(* IEC 61131-3 sources: test/Class/SafetyBaseFSoE (part 3) *)

                // get length of Name
                sd_retval := SDOReadCfgRequ ( p_SDORequestBuffer  := p_SDORequestBuffer
                                            , p_SDOResponseBuffer := p_SDOResponseBuffer
                                            , ud_Address          := ud_Address
                                            , us_Length           := 4
                                            );
                //no response
                if ( sd_retval <> 0 ) then
                  LogError("@020A (SafetyBaseFSoE::ReadSDOConfig) Config Read Error: Reading length of unsafe BDINT output name failed.");
                  return;
                end_if;

                // prepare address to get name
                ud_Address += 4;

  //              ud_ActStrLen := ud_TmpStrLen := p_SDOResponseBuffer^.ud_Data;
                ud_TmpStrLen := p_SDOResponseBuffer^.ud_Data;
                ud_ActStrLen := ud_TmpStrLen;
                ud_TmpAddress := ud_Address;

                IF p_BlockedTransferMemory = NIL THEN
                  sd_retval := -100;
                  SetSafetyState(NewState:=_MemAllocFailed);
                  RETURN;
                END_IF;

                IF ud_BlockedTransferMemorySize < (ud_TmpStrLen + 1) THEN
                  p_BlockedTransferMemory := ToStdLib.ReAlloc(mptr:=p_BlockedTransferMemory, newsize:=GetNewMemSize(ud_TmpStrLen + 1));
                  IF p_BlockedTransferMemory = NIL THEN
                    ud_BlockedTransferMemorySize := 0;
                    sd_retval := -100;
                    SetSafetyState(NewState:=_MemAllocFailed);
                    RETURN;
                  ELSE
                    ud_BlockedTransferMemorySize := GetNewMemSize(ud_TmpStrLen + 1);
                  END_IF;
                END_IF;

                ToStdLib.MemSet(dest:=p_BlockedTransferMemory, value:=0, size:=ud_BlockedTransferMemorySize);

                p_TmpBlockedData := p_BlockedTransferMemory;

                us_BlockedTransferLength := BlockedTransferLength(ud_Datalength:=ud_TmpStrLen, us_MaxBlocklength:=60);

                while us_BlockedTransferLength do

                  // get name
                  sd_retval := SDOReadCfgRequ ( p_SDORequestBuffer  := p_SDORequestBuffer
                                              , p_SDOResponseBuffer := p_SDOResponseBuffer
                                              , ud_Address          := ud_TmpAddress
                                              , us_Length           := us_BlockedTransferLength
                                              , b_UseCache          := us_BlockedTransferLength < us_DataLength_Max
                                              );
                  //no response
                  if ( sd_retval <> 0 ) then
                    LogError("@0207 (SafetyBaseFSoE::ReadSDOConfig) Config Read Error: Reading unsafe BDINT output name failed.");
                    return;
                  end_if;

                  ToStdLib.MemCpy(dest:=p_TmpBlockedData,
                                   source:=#p_SDOResponseBuffer^.ud_Data,
                                   size:=us_BlockedTransferLength);

                  p_TmpBlockedData += us_BlockedTransferLength;
                  ud_TmpAddress += us_BlockedTransferLength;
                  ud_TmpStrLen -= us_BlockedTransferLength;

                  us_BlockedTransferLength := BlockedTransferLength(ud_Datalength:=ud_TmpStrLen, us_MaxBlocklength:=60);

                end_while;

                ActBitMask := (pBitMasks + (i-1) * sizeof(BDINT))^;

                // if unsafe component not found (sd_retval <> 0), it's not problem for whole safe application

                sd_retval :=AddFastUnsafeRoutElement(pRoutTable:=#p_FastUnsafeOutputsTable,
                                                     pRoutElementsNo:=#ui_CntFastUnsafeOutputs,
                                                     ud_Address:=ud_FastUnsafe_Offset_Out,
                                                     ui_NameLen:=ud_ActStrLen$UINT,
                                                     pNameNewElement:=p_BlockedTransferMemory$^CHAR,
                                                     ActBitMask,
                                                     bWriteVar:=TRUE);

                // get offset in application memory
                ud_ActAddress += CountBits(ActBitMask) * sizeof(DINT);
                ud_FastUnsafe_Offset_Out += sizeof(DINT);

                // prepare address for next unsafe output or for number of safe inputs
                ud_Address += ud_ActStrLen;

              end_for;

              // free the bitmasks
              ToStdLib.Free(mptr:=pBitMasks);

            end_if;

          end_if; //b_IprCodeLengthAvailable = FALSE

        end_if; //b_CfgTypeV2

//*****************************************************************************
//**   UNSAFE BOOL OUTPUT VARIABLES                                          **
//*****************************************************************************

        //read number of unsafe output vars

        //send request and receive data
        sd_retval := SDOReadCfgRequ ( p_SDORequestBuffer  := p_SDORequestBuffer
                                    , p_SDOResponseBuffer := p_SDOResponseBuffer
                                    , ud_Address          := ud_Address
                                    , us_Length           := 4
                                    );

        //no response
        if ( sd_retval <> 0 ) then
          LogError("@0204 (SafetyBaseFSoE::ReadSDOConfig) Config Read Error: Reading number of unsafe bool output vars failed.");
          return;
        end_if;

        ud_CntUnsafeOutputs := p_SDOResponseBuffer^.ud_Data;

        ud_Address += 4;

        // skip the names of unsafe outputs
        for i := 1 to ud_CntUnsafeOutputs do

          // get length of Name
          sd_retval := SDOReadCfgRequ ( p_SDORequestBuffer  := p_SDORequestBuffer
                                      , p_SDOResponseBuffer := p_SDOResponseBuffer
                                      , ud_Address          := ud_Address
                                      , us_Length           := 4
                                      );
          //no response
          if ( sd_retval <> 0 ) then
            LogError("@0205 (SafetyBaseFSoE::ReadSDOConfig) Config Read Error: Reading length of unsafe bool output name failed.");
            return;
          end_if;

          // prepare address to get name
          ud_Address += 4;

//          ud_ActStrLen := ud_TmpStrLen := p_SDOResponseBuffer^.ud_Data;
          ud_TmpStrLen := p_SDOResponseBuffer^.ud_Data;
          ud_ActStrLen := ud_TmpStrLen;
          ud_TmpAddress := ud_Address;

          IF p_BlockedTransferMemory = NIL THEN
            sd_retval := -100;
            SetSafetyState(NewState:=_MemAllocFailed);
            RETURN;
          END_IF;

          IF ud_BlockedTransferMemorySize < (ud_TmpStrLen + 1) THEN
            p_BlockedTransferMemory := ToStdLib.ReAlloc(mptr:=p_BlockedTransferMemory, newsize:=GetNewMemSize(ud_TmpStrLen + 1));
            IF p_BlockedTransferMemory = NIL THEN
              ud_BlockedTransferMemorySize := 0;
              sd_retval := -100;
              SetSafetyState(NewState:=_MemAllocFailed);
              RETURN;
            ELSE
              ud_BlockedTransferMemorySize := GetNewMemSize(ud_TmpStrLen + 1);
            END_IF;
          END_IF;

          ToStdLib.MemSet(dest:=p_BlockedTransferMemory, value:=0, size:=ud_BlockedTransferMemorySize);

          p_TmpBlockedData := p_BlockedTransferMemory;

          us_BlockedTransferLength := BlockedTransferLength(ud_Datalength:=ud_TmpStrLen, us_MaxBlocklength:=60);

          while us_BlockedTransferLength do

            // get name
            sd_retval := SDOReadCfgRequ ( p_SDORequestBuffer  := p_SDORequestBuffer
                                        , p_SDOResponseBuffer := p_SDOResponseBuffer
                                        , ud_Address          := ud_TmpAddress
                                        , us_Length           := us_BlockedTransferLength
                                        , b_UseCache          := us_BlockedTransferLength < us_DataLength_Max
                                        );
            //no response
            if ( sd_retval <> 0 ) then
              LogError("0206 (SafetyBaseFSoE::ReadSDOConfig) Config Read Error: Reading unsafe bool output name failed.");
              return;
            end_if;

            ToStdLib.MemCpy(dest:=p_TmpBlockedData,
                             source:=#p_SDOResponseBuffer^.ud_Data,
                             size:=us_BlockedTransferLength);

            p_TmpBlockedData += us_BlockedTransferLength;
            ud_TmpAddress += us_BlockedTransferLength;
            ud_TmpStrLen -= us_BlockedTransferLength;

            us_BlockedTransferLength := BlockedTransferLength(ud_Datalength:=ud_TmpStrLen, us_MaxBlocklength:=60);

          end_while;

          sd_retval := AddUnsafeRoutElement(pRoutTable:=#p_UnsafeOutputsTable,
                                            pRoutElementsNo:=#ui_CntUnsafeOutputs,
                                            ud_Address:=ud_ActAddress,
                                            ui_NameLen:=ud_ActStrLen$UINT,
                                            pNameNewElement:=p_BlockedTransferMemory$^CHAR);

          // if unsafe component not found (sd_retval <> 0), it's not problem for whole safe application

          // get offset in application memory
          ud_ActAddress += 4;

          // prepare address for next unsafe output or for number of safe inputs
          ud_Address += ud_ActStrLen;

        end_for;

        // special unsafe variables (not supported by old modules)
        if b_CfgTypeV2 then

//*****************************************************************************
//**   UNSAFE BDINT OUTPUT VARIABLES                                         **
//*****************************************************************************

          //read number of unsafe BDINT output vars

          //send request and receive data
          sd_retval := SDOReadCfgRequ ( p_SDORequestBuffer  := p_SDORequestBuffer
                                      , p_SDOResponseBuffer := p_SDOResponseBuffer
                                      , ud_Address          := ud_Address
                                      , us_Length           := 4
                                      );

          //no response
          if ( sd_retval <> 0 ) then
            LogError("@0207 (SafetyBaseFSoE::ReadSDOConfig) Config Read Error: Reading number of unsafe BDINT output vars failed.");
            return;
          end_if;

          ud_CntUnsafeOutputs := p_SDOResponseBuffer^.ud_Data;

          ud_Address += 4;

          if ud_CntUnsafeOutputs then

            //SDO request for this command has 5 bytes additional data
            pBitMasks$^void := ToStdLib.Malloc(size := ud_CntUnsafeOutputs * sizeof(BDINT));

            if ( pBitMasks = NIL ) then
              sd_retval                         := -100;
              SetSafetyState(NewState:=_MemAllocFailed);
              LogError("@0208 (SafetyBaseFSoE::ReadSDOConfig) Config Read Error: Failed to allocate memory for the BDINT variable bitmasks.");
              return;
            end_if;

            // get the bitmasks for the BDINT variables
            for i := 1 to ud_CntUnsafeOutputs do

              // get bitmask
              sd_retval := SDOReadCfgRequ ( p_SDORequestBuffer  := p_SDORequestBuffer
                                          , p_SDOResponseBuffer := p_SDOResponseBuffer
                                          , ud_Address          := ud_Address
                                          , us_Length           := 4
                                          );
              //no response
              if ( sd_retval <> 0 ) then
                LogError("@0207 (SafetyBaseFSoE::ReadSDOConfig) Config Read Error: Reading bit mask of unsafe BDINT output failed.");
                return;
              end_if;

              // prepare address for the next one
              ud_Address += 4;

              // save the bitmask for adding the rout element
              (pBitMasks + (i-1) * sizeof(BDINT))^ := p_SDOResponseBuffer^.ud_Data;
            end_for;

            // skip the names of unsafe outputs
            for i := 1 to ud_CntUnsafeOutputs do

              // get length of Name
              sd_retval := SDOReadCfgRequ ( p_SDORequestBuffer  := p_SDORequestBuffer
                                          , p_SDOResponseBuffer := p_SDOResponseBuffer
                                          , ud_Address          := ud_Address
                                          , us_Length           := 4
                                          );
              //no response
              if ( sd_retval <> 0 ) then
                LogError("@020A (SafetyBaseFSoE::ReadSDOConfig) Config Read Error: Reading length of unsafe BDINT output name failed.");
                return;
              end_if;

              // prepare address to get name
              ud_Address += 4;

//              ud_ActStrLen := ud_TmpStrLen := p_SDOResponseBuffer^.ud_Data;
              ud_TmpStrLen := p_SDOResponseBuffer^.ud_Data;
              ud_ActStrLen := ud_TmpStrLen;
              ud_TmpAddress := ud_Address;

              IF p_BlockedTransferMemory = NIL THEN
                sd_retval := -100;
                SetSafetyState(NewState:=_MemAllocFailed);
                RETURN;
              END_IF;

              IF ud_BlockedTransferMemorySize < (ud_TmpStrLen + 1) THEN
                p_BlockedTransferMemory := ToStdLib.ReAlloc(mptr:=p_BlockedTransferMemory, newsize:=GetNewMemSize(ud_TmpStrLen + 1));
                IF p_BlockedTransferMemory = NIL THEN
                  ud_BlockedTransferMemorySize := 0;
                  sd_retval := -100;
                  SetSafetyState(NewState:=_MemAllocFailed);
                  RETURN;
                ELSE
                  ud_BlockedTransferMemorySize := GetNewMemSize(ud_TmpStrLen + 1);
                END_IF;
              END_IF;

              ToStdLib.MemSet(dest:=p_BlockedTransferMemory, value:=0, size:=ud_BlockedTransferMemorySize);

              p_TmpBlockedData := p_BlockedTransferMemory;

              us_BlockedTransferLength := BlockedTransferLength(ud_Datalength:=ud_TmpStrLen, us_MaxBlocklength:=60);

              while us_BlockedTransferLength do

                // get name
                sd_retval := SDOReadCfgRequ ( p_SDORequestBuffer  := p_SDORequestBuffer
                                            , p_SDOResponseBuffer := p_SDOResponseBuffer
                                            , ud_Address          := ud_TmpAddress
                                            , us_Length           := us_BlockedTransferLength
                                            , b_UseCache          := us_BlockedTransferLength < us_DataLength_Max
                                            );
                //no response
                if ( sd_retval <> 0 ) then
                  LogError("@0207 (SafetyBaseFSoE::ReadSDOConfig) Config Read Error: Reading unsafe BDINT output name failed.");
                  return;
                end_if;

                ToStdLib.MemCpy(dest:=p_TmpBlockedData,
                                 source:=#p_SDOResponseBuffer^.ud_Data,
                                 size:=us_BlockedTransferLength);

                p_TmpBlockedData += us_BlockedTransferLength;
                ud_TmpAddress += us_BlockedTransferLength;
                ud_TmpStrLen -= us_BlockedTransferLength;

                us_BlockedTransferLength := BlockedTransferLength(ud_Datalength:=ud_TmpStrLen, us_MaxBlocklength:=60);

              end_while;

              ActBitMask := (pBitMasks + (i-1) * sizeof(BDINT))^;

              sd_retval := AddUnsafeRoutElement(pRoutTable:=#p_UnsafeOutputsTable,
                                                pRoutElementsNo:=#ui_CntUnsafeOutputs,
                                                ud_Address:=ud_UnsafeBDINT_Offset,
                                                ui_NameLen:=ud_ActStrLen$UINT,
                                                pNameNewElement:=p_BlockedTransferMemory$^CHAR,
                                                ActBitMask);

              // if unsafe component not found (sd_retval <> 0), it's not problem for whole safe application

              // get offset in application memory
              ud_ActAddress += CountBits(ActBitMask) * sizeof(DINT);
              ud_UnsafeBDINT_Offset += sizeof(DINT);

              // prepare address for next unsafe output or for number of safe inputs
              ud_Address += ud_ActStrLen;

            end_for;

            // free the bitmasks
            ToStdLib.Free(mptr:=pBitMasks);
          end_if;
        end_if;

//*****************************************************************************
//**   SAFE INPUT VARIABLES                                                  **
//*****************************************************************************

        // get number of safe inputs
        sd_retval := SDOReadCfgRequ ( p_SDORequestBuffer  := p_SDORequestBuffer
                                    , p_SDOResponseBuffer := p_SDOResponseBuffer
                                    , ud_Address          := ud_Address
                                    , us_Length           := 4
                                    );

        //no response
        if ( sd_retval <> 0 ) then
          LogError("@020B (SafetyBaseFSoE::ReadSDOConfig) Config Read Error: Reading number of safe inputs failed.");
          return;
        end_if;

        //number of safe inputs
        ud_TmpCnt := p_SDOResponseBuffer^.ud_Data;

        // get offset in application memory
        ud_ActAddress += ud_TmpCnt * 4;

        //address of path length of first safe input
        ud_Address := p_SDORequestBuffer^.ud_Address + 4;

        if ud_TmpCnt then
          //read path of all safe inputs and add them to routing lists
          for i := 1 to ud_TmpCnt do

            //read path
            sd_retval := ReadModulePath ( p_SDORequestBuffer          := p_SDORequestBuffer
                                        , p_SDOResponseBuffer         := p_SDOResponseBuffer
                                        , p_ud_Address                := #ud_Address
                                        , pModule                     := pModule
                                        , p_ud_ModulePathLen_Max      := #ud_ModulePathLen_Max
                                        , p_ud_ModulePathCompLen_Max  := #ud_ModulePathCompLen_Max
                                        , us_SDOMaxDataSize           := us_DataLength_Max
                                        );

            //no response, error
            if ( sd_retval <> 0 ) then
              LogError("@020C (SafetyBaseFSoE::ReadSDOConfig) Config Read Error: Reading path of safe input failed.");
              return;
            end_if;

            // if there is a valid module path
            if pModule^.p_us_Path <> NIL then
              //add module to routing tabs
              sd_retval := AddModuleToRoutingTabs ( pModule       := pModule
                                                  , pListHeader   := pListHeader
                                                  , b_IsOptional  := TempModuleConfig.Info.IsOptional
                                                  );

              if (sd_retval <> 0 ) then
                if ( SafetyState <> _ModFromCfgNotFound ) then
                  LogError("@020D (SafetyBaseFSoE::ReadSDOConfig) Config Read Error: Failed to add safe input module to routing tabs.");
                  return;
                end_if;
              end_if;
            end_if;

            if b_IsFSoE then
              // lower 2 Bytes: Index in connection list, upper 2 Bytes: Bit-Offset of the value inside the process data (not the FSoE frame)
              ud_Address += 4;
            else
              //address of path length = last address + 2 * 4 bytes ( RemoteIndex + MaxAge)
              ud_Address += 8;
            end_if;
          end_for;
        end_if;

        if b_CfgTypeV3 then

//*****************************************************************************
//**   SAFE DINT INPUT VARIABLES                                             **
//*****************************************************************************

          // get number of safe DINT inputs
          sd_retval := SDOReadCfgRequ ( p_SDORequestBuffer  := p_SDORequestBuffer
                                      , p_SDOResponseBuffer := p_SDOResponseBuffer
                                      , ud_Address          := ud_Address
                                      , us_Length           := 4
                                      );

          //no response
          if ( sd_retval <> 0 ) then
            LogError("@020E (SafetyBaseFSoE::ReadSDOConfig) Config Read Error: Reading number of safe DINT inputs failed.");
            return;
          end_if;

          //number of safe inputs
          ud_TmpCnt := p_SDOResponseBuffer^.ud_Data;

          // get offset in application memory
          ud_ActAddress += ud_TmpCnt * 8;

          //address of path length of first safe input
          ud_Address := p_SDORequestBuffer^.ud_Address + 4;

          //read path of all safe inputs and add them to routing lists
          for i := 1 to ud_TmpCnt do

            //read path
            sd_retval := ReadModulePath ( p_SDORequestBuffer          := p_SDORequestBuffer
                                        , p_SDOResponseBuffer         := p_SDOResponseBuffer
                                        , p_ud_Address                := #ud_Address
                                        , pModule                     := pModule
                                        , p_ud_ModulePathLen_Max      := #ud_ModulePathLen_Max
                                        , p_ud_ModulePathCompLen_Max  := #ud_ModulePathCompLen_Max
                                        , us_SDOMaxDataSize           := us_DataLength_Max
                                        );

            //no response, error
            if ( sd_retval <> 0 ) then
              LogError("@020F (SafetyBaseFSoE::ReadSDOConfig) Config Read Error: Reading path of safe DINT input failed.");
              return;
            end_if;

            // if there is a valid module path
            if pModule^.p_us_Path <> NIL then
              //add module to routing tabs
              sd_retval := AddModuleToRoutingTabs ( pModule       := pModule
                                                  , pListHeader   := pListHeader
                                                  , b_IsOptional  := TempModuleConfig.Info.IsOptional
                                                  );

              if (sd_retval <> 0 ) then
                if ( SafetyState <> _ModFromCfgNotFound ) then
                  LogError("@0210 (SafetyBaseFSoE::ReadSDOConfig) Config Read Error: Failed to add safe DINT input module to routing tabs.");
                  return;
                end_if;
              end_if;
            end_if;

            if b_IsFSoE then
              // lower 2 Bytes: Index in connection list, upper 2 Bytes: Bit-Offset of the value inside the process data (not the FSoE frame)
              ud_Address += 4;
            else
              //address of path length = last address + 2 * 4 bytes ( RemoteIndex + MaxAge)
              ud_Address += 8;
            end_if;
          end_for;
        end_if;

        // only available at new modules
        if b_CfgTypeV2 then

//*****************************************************************************
//**   SAFE INTERFACE INPUT VARIABLES                                        **
//*****************************************************************************

          // get number of safe interface input vars

          //send request and receive data
          sd_retval := SDOReadCfgRequ ( p_SDORequestBuffer  := p_SDORequestBuffer
                                      , p_SDOResponseBuffer := p_SDOResponseBuffer
                                      , ud_Address          := ud_Address
                                      , us_Length           := 4
                                      );

          //no response
          if ( sd_retval <> 0 ) then
            LogError("@0211 (SafetyBaseFSoE::ReadSDOConfig) Config Read Error: Reading number of safe interface input variables failed.");
            return;
          end_if;

          // skip the number
          ud_Address += 4;

          //number of safe inputs
          ud_TmpCnt := p_SDOResponseBuffer^.ud_Data;

          // get offset in application memory
          ud_ActAddress += ud_TmpCnt * 4;

          if ud_TmpCnt then

            for i := 0 to (ud_TmpCnt-1) do
              // get length of the uncompressed path

              //send request and receive data
              sd_retval := SDOReadCfgRequ ( p_SDORequestBuffer  := p_SDORequestBuffer
                                          , p_SDOResponseBuffer := p_SDOResponseBuffer
                                          , ud_Address          := ud_Address
                                          , us_Length           := 4
                                          );

              //no response
              if ( sd_retval <> 0 ) then
                LogError("@0212 (SafetyBaseFSoE::ReadSDOConfig) Config Read Error: Reading length of uncompressed interface topology path failed.");
                return;
              end_if;

              // skip length of top path
              ud_Address += 4;

              // skip top path
              ud_Address += p_SDOResponseBuffer^.ud_Data;

              // read length of compressed topology path

              //send request and receive data
              sd_retval := SDOReadCfgRequ ( p_SDORequestBuffer  := p_SDORequestBuffer
                                          , p_SDOResponseBuffer := p_SDOResponseBuffer
                                          , ud_Address          := ud_Address
                                          , us_Length           := 4
                                          );

              //no response
              if ( sd_retval <> 0 ) then
                LogError("@0279 (SafetyBaseFSoE::ReadSDOConfig) Config Read Error: Reading length of compressed interface topology path failed.");
                return;
              end_if;

              // skip length of compressed top path and compressed top path
              ud_Address += 4 + p_SDOResponseBuffer^.ud_Data;

              if b_IsFSoE then
                // lower 2 Bytes: Index in connection list, upper 2 Bytes: Bit-Offset of the value inside the process data (not the FSoE frame)
                ud_Address += 4;
              else
                //address of path length = last address + 2 * 4 bytes ( RemoteIndex + MaxAge)
                ud_Address += 8;
              end_if;
            end_for;
          end_if;

(*
 4 Byte Anzahl
 4 Byte Länge vom Pfad, Pfad (vorne Pfad ":" dann CRC für da Interface dann bis auf 4 Byte aufgefüllt)
 4 Byte Länge vom komprimierten Pfad, komprimierter Pfad (vorne Pfad ":" dann CRC für da Interface dann bis auf 4 Byte aufgefüllt)
 4 Byte RemoteIndex
 4 Byte Maximales Alter
*)

        end_if;

        // only available at new containers
        if b_CfgTypeV3 then

//*****************************************************************************
//**   SAFE DINT INTERFACE INPUT VARIABLES                                   **
//*****************************************************************************

          // get number of safe DINT interface input vars

          //send request and receive data
          sd_retval := SDOReadCfgRequ ( p_SDORequestBuffer  := p_SDORequestBuffer
                                      , p_SDOResponseBuffer := p_SDOResponseBuffer
                                      , ud_Address          := ud_Address
                                      , us_Length           := 4
                                      );

          //no response
          if ( sd_retval <> 0 ) then
            LogError("@0213 (SafetyBaseFSoE::ReadSDOConfig) Config Read Error: Reading number of safe DINT interface input variables failed.");
            return;
          end_if;

          // skip the number
          ud_Address += 4;

          //number of safe inputs
          ud_TmpCnt := p_SDOResponseBuffer^.ud_Data;

          // get offset in application memory
          ud_ActAddress += ud_TmpCnt * 8;

          if ud_TmpCnt then

            for i := 0 to (ud_TmpCnt-1) do
              // get length of the uncompressed path

              //send request and receive data
              sd_retval := SDOReadCfgRequ ( p_SDORequestBuffer  := p_SDORequestBuffer
                                          , p_SDOResponseBuffer := p_SDOResponseBuffer
                                          , ud_Address          := ud_Address
                                          , us_Length           := 4
                                          );

              //no response
              if ( sd_retval <> 0 ) then
                LogError("@0214 (SafetyBaseFSoE::ReadSDOConfig) Config Read Error: Reading length of uncompressed interface topology path failed at safe DINT input variables.");
                return;
              end_if;

              // skip length of top path
              ud_Address += 4;

              // skip top path
              ud_Address += p_SDOResponseBuffer^.ud_Data;

              // read length of compressed topology path

              //send request and receive data
              sd_retval := SDOReadCfgRequ ( p_SDORequestBuffer  := p_SDORequestBuffer
                                          , p_SDOResponseBuffer := p_SDOResponseBuffer
                                          , ud_Address          := ud_Address
                                          , us_Length           := 4
                                          );

              //no response
              if ( sd_retval <> 0 ) then
                LogError("@0215 (SafetyBaseFSoE::ReadSDOConfig) Config Read Error: Reading length of compressed interface topology path failed at safe DINT input variables.");
                return;
              end_if;

              // skip length of compressed top path and compressed top path
              ud_Address += 4 + p_SDOResponseBuffer^.ud_Data;

              if b_IsFSoE then
                // lower 2 Bytes: Index in connection list, upper 2 Bytes: Bit-Offset of the value inside the process data (not the FSoE frame)
                ud_Address += 4;
              else
                //address of path length = last address + 2 * 4 bytes ( RemoteIndex + MaxAge)
                ud_Address += 8;
              end_if;
            end_for;
          end_if;

(*
 4 Byte Anzahl
 4 Byte Länge vom Pfad, Pfad (vorne Pfad ":" dann CRC für da Interface dann bis auf 4 Byte aufgefüllt)
 4 Byte Länge vom komprimierten Pfad, komprimierter Pfad (vorne Pfad ":" dann CRC für da Interface dann bis auf 4 Byte aufgefüllt)
 4 Byte RemoteIndex
 4 Byte Maximales Alter
*)

        end_if;

//*****************************************************************************
//**   FAST UNSAFE INPUT VARIABLES                                           **
//*****************************************************************************

        // only available at new modules
        if b_CfgTypeV2 then

          if b_IprCodeLengthAvailable = FALSE then
            // get number of fast unsafe intput vars

            //send request and receive data
            sd_retval := SDOReadCfgRequ ( p_SDORequestBuffer  := p_SDORequestBuffer
                                        , p_SDOResponseBuffer := p_SDOResponseBuffer
                                        , ud_Address          := ud_Address
                                        , us_Length           := 4
                                        );

            //no response
            if ( sd_retval <> 0 ) then
              LogError("@0216 (SafetyBaseFSoE::ReadSDOConfig) Config Read Error: Reading number of fast unsafe intput vars failed.");
              return;
            end_if;

            ud_Address += 4;

            // get offset in application memory
            ud_ActAddress += p_SDOResponseBuffer^.ud_Data * 4;
            // if it's our own path, remember the fast unsafe settings
            if (PathOfThisCPU[0]$UINT = (pListHeader^.p_us_Path$^UINT)^) & (ToStdLib.MemCmp(#PathOfThisCPU[0], pListHeader^.p_us_Path, PathOfThisCPU[0]$UINT + 2) = 0) then
              if (p_SDOResponseBuffer^.ud_Data <> 0) then
                if ActivateFastUnsafeIOs then
                  b_FastUnsafeInputsActive := TRUE;
                else
                  // error => can't go on like this
                  LogError("@0202 (SafetyBaseFSoE::ReadSDOConfig) Number or size of module accesses increased with new safety project!");
                  LogError("@0203 (SafetyBaseFSoE::ReadSDOConfig) => Can't continue, because the new data is not covered by the actual accesses! Restart Application!");

                  b_NeedApplicationRestart := TRUE;
                end_if;
              end_if;
            end_if;
          else  //b_IprCodeLengthAvailable = FALSE

//*****************************************************************************
//**   Fast UNSAFE BOOL INPUT VARIABLES     SCP211                           **
//*****************************************************************************

            // here we go for unsafe bool input vars

            // get number of unsafe input vars
            sd_retval := SDOReadCfgRequ ( p_SDORequestBuffer  := p_SDORequestBuffer
                                        , p_SDOResponseBuffer := p_SDOResponseBuffer
                                        , ud_Address          := ud_Address
                                        , us_Length           := 4
                                        );

            //no response
            if ( sd_retval <> 0 ) then
              LogError("@0217 (SafetyBaseFSoE::ReadSDOConfig) Config Read Error: Failed to read number of unsafe input vars.");
              return;
            end_if;

            ud_CntFastUnsafeInputs:= p_SDOResponseBuffer^.ud_Data;

            ud_Address += 4;

            // skip the names of unsafe inputs
            for i := 1 to ud_CntFastUnsafeInputs do

              // get length of Name
              sd_retval := SDOReadCfgRequ ( p_SDORequestBuffer  := p_SDORequestBuffer
                                          , p_SDOResponseBuffer := p_SDOResponseBuffer
                                          , ud_Address          := ud_Address
                                          , us_Length           := 4
                                          );
              //no response
              if ( sd_retval <> 0 ) then
                LogError("@0218 (SafetyBaseFSoE::ReadSDOConfig) Config Read Error: Reading length of unsafe input name failed.");
                return;
              end_if;

              // prepare address to get name
              ud_Address += 4;

    //          ud_ActStrLen := ud_TmpStrLen := p_SDOResponseBuffer^.ud_Data;
              ud_TmpStrLen := p_SDOResponseBuffer^.ud_Data;
              ud_ActStrLen := ud_TmpStrLen;
              ud_TmpAddress := ud_Address;

              IF p_BlockedTransferMemory = NIL THEN
                sd_retval := -100;
                SetSafetyState(NewState:=_MemAllocFailed);
                RETURN;
              END_IF;

              IF ud_BlockedTransferMemorySize < (ud_TmpStrLen + 1) THEN
                p_BlockedTransferMemory := ToStdLib.ReAlloc(mptr:=p_BlockedTransferMemory, newsize:=GetNewMemSize(ud_TmpStrLen + 1));
                IF p_BlockedTransferMemory = NIL THEN
                  ud_BlockedTransferMemorySize := 0;
                  sd_retval := -100;
                  SetSafetyState(NewState:=_MemAllocFailed);
                  RETURN;
                ELSE
                  ud_BlockedTransferMemorySize := GetNewMemSize(ud_TmpStrLen + 1);
                END_IF;
              END_IF;

              ToStdLib.MemSet(dest:=p_BlockedTransferMemory, value:=0, size:=ud_BlockedTransferMemorySize);

              p_TmpBlockedData := p_BlockedTransferMemory;

              us_BlockedTransferLength := BlockedTransferLength(ud_Datalength:=ud_TmpStrLen, us_MaxBlocklength:=60);

              while us_BlockedTransferLength do

                // get name
                sd_retval := SDOReadCfgRequ ( p_SDORequestBuffer  := p_SDORequestBuffer
                                            , p_SDOResponseBuffer := p_SDOResponseBuffer
                                            , ud_Address          := ud_TmpAddress
                                            , us_Length           := us_BlockedTransferLength
                                            , b_UseCache          := us_BlockedTransferLength < us_DataLength_Max
                                            );
                //no response
                if ( sd_retval <> 0 ) then
                  LogError("@0219 (SafetyBaseFSoE::ReadSDOConfig) Config Read Error: Reading unsafe input name failed.");
                  return;
                end_if;

                ToStdLib.MemCpy(dest:=p_TmpBlockedData,
                                 source:=#p_SDOResponseBuffer^.ud_Data,
                                 size:=us_BlockedTransferLength);

                p_TmpBlockedData += us_BlockedTransferLength;
                ud_TmpAddress += us_BlockedTransferLength;
                ud_TmpStrLen -= us_BlockedTransferLength;

                us_BlockedTransferLength := BlockedTransferLength(ud_Datalength:=ud_TmpStrLen, us_MaxBlocklength:=60);

              end_while;

              sd_retval := AddFastUnsafeRoutElement(pRoutTable:=#p_FastUnsafeInputsTable,
                                                    pRoutElementsNo:=#ui_CntFastUnsafeInputs,
                                                    ud_Address:=ud_FastUnsafe_Offset_In,
                                                    ui_NameLen:=ud_ActStrLen$UINT,
                                                    pNameNewElement:=p_BlockedTransferMemory$^CHAR,
                                                    bWriteVar:=FALSE);

              // if unsafe component not found (sd_retval <> 0), it's not problem for whole safe application
              // get offset in application memory
              ud_ActAddress += 4;
              ud_FastUnsafe_Offset_In += sizeof(DINT);

              // prepare address for next unsafe input
              ud_Address += ud_ActStrLen;

            end_for;

//*****************************************************************************
//**  FAST UNSAFE BDINT INPUT VARIABLES       SCP211                         **
//*****************************************************************************

            // here we go for unsafe BDINT input vars

            // get number of unsafe input vars
            sd_retval := SDOReadCfgRequ ( p_SDORequestBuffer  := p_SDORequestBuffer
                                        , p_SDOResponseBuffer := p_SDOResponseBuffer
                                        , ud_Address          := ud_Address
                                        , us_Length           := 4
                                        );

            //no response
            if ( sd_retval <> 0 ) then
              LogError("@021A (SafetyBaseFSoE::ReadSDOConfig) Config Read Error: Failed to read number of unsafe BDINT input vars.");
              return;
            end_if;

            ud_CntFastUnsafeInputs := p_SDOResponseBuffer^.ud_Data;

            ud_Address += 4;

            if ud_CntFastUnsafeInputs then

              //SDO request for this command has 5 bytes additional data
              pBitMasks$^void := ToStdLib.Malloc(size := ud_CntFastUnsafeInputs * sizeof(BDINT));

              if ( pBitMasks = NIL ) then
                sd_retval                         := -100;
                SetSafetyState(NewState:=_MemAllocFailed);
                LogError("@021B (SafetyBaseFSoE::ReadSDOConfig) Config Read Error: Failed to allocate memory for the BDINT variable bitmasks.");
                return;
              end_if;

              // get the bitmasks for the BDINT variables
              for i := 1 to ud_CntFastUnsafeInputs do

                // get bitmask
                sd_retval := SDOReadCfgRequ ( p_SDORequestBuffer  := p_SDORequestBuffer
                                            , p_SDOResponseBuffer := p_SDOResponseBuffer
                                            , ud_Address          := ud_Address
                                            , us_Length           := 4
                                            );
                //no response
                if ( sd_retval <> 0 ) then
                  LogError("021C (SafetyBaseFSoE::ReadSDOConfig) Config Read Error: Reading bit mask of unsafe BDINT input failed.");
                  return;
                end_if;

                // prepare address for the next one
                ud_Address += 4;

                // save the bitmask for adding the rout element
                (pBitMasks + (i-1) * sizeof(BDINT))^ := p_SDOResponseBuffer^.ud_Data;
              end_for;

              // get the names of unsafe inputs
              for i := 1 to ud_CntFastUnsafeInputs do

                // get length of Name
                sd_retval := SDOReadCfgRequ ( p_SDORequestBuffer  := p_SDORequestBuffer
                                            , p_SDOResponseBuffer := p_SDOResponseBuffer
                                            , ud_Address          := ud_Address
                                            , us_Length           := 4
                                            );
                //no response
                if ( sd_retval <> 0 ) then
                  LogError("@021D (SafetyBaseFSoE::ReadSDOConfig) Config Read Error: Reading length of unsafe BDINT input name failed.");
                  return;
                end_if;

                // prepare address to get name
                ud_Address += 4;

  //              ud_ActStrLen := ud_TmpStrLen := p_SDOResponseBuffer^.ud_Data;
                ud_TmpStrLen := p_SDOResponseBuffer^.ud_Data;
                ud_ActStrLen := ud_TmpStrLen;
                ud_TmpAddress := ud_Address;

                IF p_BlockedTransferMemory = NIL THEN
                  sd_retval := -100;
                  SetSafetyState(NewState:=_MemAllocFailed);
                  RETURN;
                END_IF;

                IF ud_BlockedTransferMemorySize < (ud_TmpStrLen + 1) THEN
                  p_BlockedTransferMemory := ToStdLib.ReAlloc(mptr:=p_BlockedTransferMemory, newsize:=GetNewMemSize(ud_TmpStrLen + 1));
                  IF p_BlockedTransferMemory = NIL THEN
                    ud_BlockedTransferMemorySize := 0;
                    sd_retval := -100;
                    SetSafetyState(NewState:=_MemAllocFailed);
                    RETURN;
                  ELSE
                    ud_BlockedTransferMemorySize := GetNewMemSize(ud_TmpStrLen + 1);
                  END_IF;
                END_IF;

                ToStdLib.MemSet(dest:=p_BlockedTransferMemory, value:=0, size:=ud_BlockedTransferMemorySize);

                p_TmpBlockedData := p_BlockedTransferMemory;

                us_BlockedTransferLength := BlockedTransferLength(ud_Datalength:=ud_TmpStrLen, us_MaxBlocklength:=60);

                while us_BlockedTransferLength do

                  // get name
                  sd_retval := SDOReadCfgRequ ( p_SDORequestBuffer  := p_SDORequestBuffer
                                              , p_SDOResponseBuffer := p_SDOResponseBuffer
                                              , ud_Address          := ud_TmpAddress
                                              , us_Length           := us_BlockedTransferLength
                                              , b_UseCache          := us_BlockedTransferLength < us_DataLength_Max
                                              );
                  //no response
                  if ( sd_retval <> 0 ) then
                    LogError("@021E (SafetyBaseFSoE::ReadSDOConfig) Config Read Error: Reading unsafe BDINT input name failed.");
                    return;
                  end_if;

                  ToStdLib.MemCpy(dest:=p_TmpBlockedData,
                                   source:=#p_SDOResponseBuffer^.ud_Data,
                                   size:=us_BlockedTransferLength);

                  p_TmpBlockedData += us_BlockedTransferLength;
                  ud_TmpAddress += us_BlockedTransferLength;
                  ud_TmpStrLen -= us_BlockedTransferLength;

                  us_BlockedTransferLength := BlockedTransferLength(ud_Datalength:=ud_TmpStrLen, us_MaxBlocklength:=60);

                end_while;

                ActBitMask := (pBitMasks + (i-1) * sizeof(BDINT))^;

                sd_retval := AddFastUnsafeRoutElement(pRoutTable:=#p_FastUnsafeInputsTable,
                                                      pRoutElementsNo:=#ui_CntFastUnsafeInputs,
                                                      ud_Address:=ud_FastUnsafe_Offset_In,
                                                      ui_NameLen:=ud_ActStrLen$UINT,
                                                      pNameNewElement:=p_BlockedTransferMemory$^CHAR,
                                                      BitMask:=ActBitMask,
                                                      bWriteVar:= FALSE);

                // if unsafe component not found (sd_retval <> 0), it's not problem for whole safe application

                // get offset in application memory
                ud_ActAddress += CountBits(ActBitMask) * sizeof(DINT);
                ud_FastUnsafe_Offset_In += sizeof(DINT);

                // prepare address for next unsafe output or for number of constants
                ud_Address += ud_ActStrLen;

              end_for;

              // free the bitmasks
              ToStdLib.Free(mptr:=pBitMasks);

            end_if;
        end_if;
      end_if; //b_CfgTypeV2

//*****************************************************************************
//**   UNSAFE BOOL INPUT VARIABLES                                           **
//*****************************************************************************

        // here we go for unsafe bool input vars

        // get number of unsafe input vars
        sd_retval := SDOReadCfgRequ ( p_SDORequestBuffer  := p_SDORequestBuffer
                                    , p_SDOResponseBuffer := p_SDOResponseBuffer
                                    , ud_Address          := ud_Address
                                    , us_Length           := 4
                                    );

        //no response
        if ( sd_retval <> 0 ) then
          LogError("@0217 (SafetyBaseFSoE::ReadSDOConfig) Config Read Error: Failed to read number of unsafe input vars.");
          return;
        end_if;

        ud_CntUnsafeInputs := p_SDOResponseBuffer^.ud_Data;

        ud_Address += 4;

        // skip the names of unsafe inputs
        for i := 1 to ud_CntUnsafeInputs do

          // get length of Name
          sd_retval := SDOReadCfgRequ ( p_SDORequestBuffer  := p_SDORequestBuffer
                                      , p_SDOResponseBuffer := p_SDOResponseBuffer
                                      , ud_Address          := ud_Address
                                      , us_Length           := 4
                                      );
          //no response
          if ( sd_retval <> 0 ) then
            LogError("@0218 (SafetyBaseFSoE::ReadSDOConfig) Config Read Error: Reading length of unsafe input name failed.");
            return;
          end_if;

          // prepare address to get name
          ud_Address += 4;

//          ud_ActStrLen := ud_TmpStrLen := p_SDOResponseBuffer^.ud_Data;
          ud_TmpStrLen := p_SDOResponseBuffer^.ud_Data;
          ud_ActStrLen := ud_TmpStrLen;
          ud_TmpAddress := ud_Address;

          IF p_BlockedTransferMemory = NIL THEN
            sd_retval := -100;
            SetSafetyState(NewState:=_MemAllocFailed);
            RETURN;
          END_IF;

          IF ud_BlockedTransferMemorySize < (ud_TmpStrLen + 1) THEN
            p_BlockedTransferMemory := ToStdLib.ReAlloc(mptr:=p_BlockedTransferMemory, newsize:=GetNewMemSize(ud_TmpStrLen + 1));
            IF p_BlockedTransferMemory = NIL THEN
              ud_BlockedTransferMemorySize := 0;
              sd_retval := -100;
              SetSafetyState(NewState:=_MemAllocFailed);
              RETURN;
            ELSE
              ud_BlockedTransferMemorySize := GetNewMemSize(ud_TmpStrLen + 1);
            END_IF;
          END_IF;

          ToStdLib.MemSet(dest:=p_BlockedTransferMemory, value:=0, size:=ud_BlockedTransferMemorySize);

          p_TmpBlockedData := p_BlockedTransferMemory;

          us_BlockedTransferLength := BlockedTransferLength(ud_Datalength:=ud_TmpStrLen, us_MaxBlocklength:=60);

          while us_BlockedTransferLength do

            // get name
            sd_retval := SDOReadCfgRequ ( p_SDORequestBuffer  := p_SDORequestBuffer
                                        , p_SDOResponseBuffer := p_SDOResponseBuffer
                                        , ud_Address          := ud_TmpAddress
                                        , us_Length           := us_BlockedTransferLength
                                        , b_UseCache          := us_BlockedTransferLength < us_DataLength_Max
                                        );
            //no response
            if ( sd_retval <> 0 ) then
              LogError("@0219 (SafetyBaseFSoE::ReadSDOConfig) Config Read Error: Reading unsafe input name failed.");
              return;
            end_if;

            ToStdLib.MemCpy(dest:=p_TmpBlockedData,
                             source:=#p_SDOResponseBuffer^.ud_Data,
                             size:=us_BlockedTransferLength);

            p_TmpBlockedData += us_BlockedTransferLength;
            ud_TmpAddress += us_BlockedTransferLength;
            ud_TmpStrLen -= us_BlockedTransferLength;

            us_BlockedTransferLength := BlockedTransferLength(ud_Datalength:=ud_TmpStrLen, us_MaxBlocklength:=60);

          end_while;

          sd_retval := AddUnsafeRoutElement(pRoutTable:=#p_UnsafeInputsTable,
                                            pRoutElementsNo:=#ui_CntUnsafeInputs,
                                            ud_Address:=ud_ActAddress,
                                            ui_NameLen:=ud_ActStrLen$UINT,
                                            pNameNewElement:=p_BlockedTransferMemory$^CHAR);

          // if unsafe component not found (sd_retval <> 0), it's not problem for whole safe application

          // get offset in application memory
          ud_ActAddress += 4;

          // prepare address for next unsafe input
          ud_Address += ud_ActStrLen;

        end_for;

        // only available at new modules
        if b_CfgTypeV2 then

//*****************************************************************************
//**   UNSAFE BDINT INPUT VARIABLES                                          **
//*****************************************************************************

          // here we go for unsafe BDINT input vars

          // get number of unsafe input vars
          sd_retval := SDOReadCfgRequ ( p_SDORequestBuffer  := p_SDORequestBuffer
                                      , p_SDOResponseBuffer := p_SDOResponseBuffer
                                      , ud_Address          := ud_Address
                                      , us_Length           := 4
                                      );

          //no response
          if ( sd_retval <> 0 ) then
            LogError("@021A (SafetyBaseFSoE::ReadSDOConfig) Config Read Error: Failed to read number of unsafe BDINT input vars.");
            return;
          end_if;

          ud_CntUnsafeInputs := p_SDOResponseBuffer^.ud_Data;

          ud_Address += 4;

          if ud_CntUnsafeInputs then

            //SDO request for this command has 5 bytes additional data
            pBitMasks$^void := ToStdLib.Malloc(size := ud_CntUnsafeInputs * sizeof(BDINT));

            if ( pBitMasks = NIL ) then
              sd_retval                         := -100;
              SetSafetyState(NewState:=_MemAllocFailed);
              LogError("@021B (SafetyBaseFSoE::ReadSDOConfig) Config Read Error: Failed to allocate memory for the BDINT variable bitmasks.");
              return;
            end_if;

            // get the bitmasks for the BDINT variables
            for i := 1 to ud_CntUnsafeInputs do

              // get bitmask
              sd_retval := SDOReadCfgRequ ( p_SDORequestBuffer  := p_SDORequestBuffer
                                          , p_SDOResponseBuffer := p_SDOResponseBuffer
                                          , ud_Address          := ud_Address
                                          , us_Length           := 4
                                          );
              //no response
              if ( sd_retval <> 0 ) then
                LogError("021C (SafetyBaseFSoE::ReadSDOConfig) Config Read Error: Reading bit mask of unsafe BDINT input failed.");
                return;
              end_if;

              // prepare address for the next one
              ud_Address += 4;

              // save the bitmask for adding the rout element
              (pBitMasks + (i-1) * sizeof(BDINT))^ := p_SDOResponseBuffer^.ud_Data;
            end_for;

            // get the names of unsafe inputs
            for i := 1 to ud_CntUnsafeInputs do

              // get length of Name
              sd_retval := SDOReadCfgRequ ( p_SDORequestBuffer  := p_SDORequestBuffer
                                          , p_SDOResponseBuffer := p_SDOResponseBuffer
                                          , ud_Address          := ud_Address
                                          , us_Length           := 4
                                          );
              //no response
              if ( sd_retval <> 0 ) then
                LogError("@021D (SafetyBaseFSoE::ReadSDOConfig) Config Read Error: Reading length of unsafe BDINT input name failed.");
                return;
              end_if;

              // prepare address to get name
              ud_Address += 4;

//              ud_ActStrLen := ud_TmpStrLen := p_SDOResponseBuffer^.ud_Data;
              ud_TmpStrLen := p_SDOResponseBuffer^.ud_Data;
              ud_ActStrLen := ud_TmpStrLen;
              ud_TmpAddress := ud_Address;

              IF p_BlockedTransferMemory = NIL THEN
                sd_retval := -100;
                SetSafetyState(NewState:=_MemAllocFailed);
                RETURN;
              END_IF;

              IF ud_BlockedTransferMemorySize < (ud_TmpStrLen + 1) THEN
                p_BlockedTransferMemory := ToStdLib.ReAlloc(mptr:=p_BlockedTransferMemory, newsize:=GetNewMemSize(ud_TmpStrLen + 1));
                IF p_BlockedTransferMemory = NIL THEN
                  ud_BlockedTransferMemorySize := 0;
                  sd_retval := -100;
                  SetSafetyState(NewState:=_MemAllocFailed);
                  RETURN;
                ELSE
                  ud_BlockedTransferMemorySize := GetNewMemSize(ud_TmpStrLen + 1);
                END_IF;
              END_IF;

              ToStdLib.MemSet(dest:=p_BlockedTransferMemory, value:=0, size:=ud_BlockedTransferMemorySize);

              p_TmpBlockedData := p_BlockedTransferMemory;

              us_BlockedTransferLength := BlockedTransferLength(ud_Datalength:=ud_TmpStrLen, us_MaxBlocklength:=60);

              while us_BlockedTransferLength do

                // get name
                sd_retval := SDOReadCfgRequ ( p_SDORequestBuffer  := p_SDORequestBuffer
                                            , p_SDOResponseBuffer := p_SDOResponseBuffer
                                            , ud_Address          := ud_TmpAddress
                                            , us_Length           := us_BlockedTransferLength
                                            , b_UseCache          := us_BlockedTransferLength < us_DataLength_Max
                                            );
                //no response
                if ( sd_retval <> 0 ) then
                  LogError("@021E (SafetyBaseFSoE::ReadSDOConfig) Config Read Error: Reading unsafe BDINT input name failed.");
                  return;
                end_if;

                ToStdLib.MemCpy(dest:=p_TmpBlockedData,
                                 source:=#p_SDOResponseBuffer^.ud_Data,
                                 size:=us_BlockedTransferLength);

                p_TmpBlockedData += us_BlockedTransferLength;
                ud_TmpAddress += us_BlockedTransferLength;
                ud_TmpStrLen -= us_BlockedTransferLength;

                us_BlockedTransferLength := BlockedTransferLength(ud_Datalength:=ud_TmpStrLen, us_MaxBlocklength:=60);

              end_while;

              ActBitMask := (pBitMasks + (i-1) * sizeof(BDINT))^;

              sd_retval := AddUnsafeRoutElement(pRoutTable:=#p_UnsafeInputsTable,
                                                pRoutElementsNo:=#ui_CntUnsafeInputs,
                                                ud_Address:=ud_UnsafeBDINT_Offset,
                                                ui_NameLen:=ud_ActStrLen$UINT,
                                                pNameNewElement:=p_BlockedTransferMemory$^CHAR,
                                                ActBitMask);

              // if unsafe component not found (sd_retval <> 0), it's not problem for whole safe application

              // get offset in application memory
              ud_ActAddress += CountBits(ActBitMask) * sizeof(DINT);
              ud_UnsafeBDINT_Offset += sizeof(DINT);

              // prepare address for next unsafe output or for number of constants
              ud_Address += ud_ActStrLen;

            end_for;

            // free the bitmasks
            ToStdLib.Free(mptr:=pBitMasks);
          end_if;

//*****************************************************************************
//**   CONSTANTS                                                             **
//*****************************************************************************

          // constants

          //send request and receive data
          sd_retval := SDOReadCfgRequ ( p_SDORequestBuffer  := p_SDORequestBuffer
                                      , p_SDOResponseBuffer := p_SDOResponseBuffer
                                      , ud_Address          := ud_Address
                                      , us_Length           := 4
                                      );

          //no response
          if ( sd_retval <> 0 ) then
            LogError("@021F (SafetyBaseFSoE::ReadSDOConfig) Config Read Error: Reading number of constants failed.");
            return;
          end_if;

          // skip number of constants
          ud_Address += 4;

          // skip constants
          ud_Address += p_SDOResponseBuffer^.ud_Data * 4;

          if b_CfgTypeV3 then

//*****************************************************************************
//**   SAFE DINT CONSTANTS                                                   **
//*****************************************************************************

            // constants

            //send request and receive data
            sd_retval := SDOReadCfgRequ ( p_SDORequestBuffer  := p_SDORequestBuffer
                                        , p_SDOResponseBuffer := p_SDOResponseBuffer
                                        , ud_Address          := ud_Address
                                        , us_Length           := 4
                                        );

            //no response
            if ( sd_retval <> 0 ) then
              LogError("@0220 (SafetyBaseFSoE::ReadSDOConfig) Config Read Error: Reading number of safe DINT constants failed.");
              return;
            end_if;

            // skip number of safe dint constants
            ud_Address += 4;

            // skip constants (4 byte per safe DINT constant)
            ud_Address += p_SDOResponseBuffer^.ud_Data * 4;

          end_if;

//*****************************************************************************
//**   LOCAL OUTPUTS                                                         **
//*****************************************************************************

          // local outputs
          //send request and receive data
          sd_retval := SDOReadCfgRequ ( p_SDORequestBuffer  := p_SDORequestBuffer
                                      , p_SDOResponseBuffer := p_SDOResponseBuffer
                                      , ud_Address          := ud_Address
                                      , us_Length           := 4
                                      );

          //no response
          if ( sd_retval <> 0 ) then
            LogError("@0221 (SafetyBaseFSoE::ReadSDOConfig) Config Read Error: Reading number of local outputs failed.");
            return;
          end_if;

          // skip number of local outputs
          ud_Address += 4;

          // skip local outputs
          //++pr
          // only available at new modules
          if b_CfgTypeV2 then
            ud_Address += p_SDOResponseBuffer^.ud_Data * 8; // Used-Flag, Modulkennung(SDIAS)
          else
            ud_Address += p_SDOResponseBuffer^.ud_Data * 4; // Used-Flag
          end_if;

          if b_CfgTypeV3 then

//*****************************************************************************
//**   LOCAL DINT OUTPUTS                                                    **
//*****************************************************************************

            // local outputs
            //send request and receive data
            sd_retval := SDOReadCfgRequ ( p_SDORequestBuffer  := p_SDORequestBuffer
                                        , p_SDOResponseBuffer := p_SDOResponseBuffer
                                        , ud_Address          := ud_Address
                                        , us_Length           := 4
                                        );

            //no response
            if ( sd_retval <> 0 ) then
              LogError("@0222 (SafetyBaseFSoE::ReadSDOConfig) Config Read Error: Reading number of local outputs failed.");
              return;
            end_if;

            // skip number of local outputs
            ud_Address += 4;

            // skip local outputs
            //++pr
            // only available at new modules
            if b_CfgTypeV2 then
              ud_Address += p_SDOResponseBuffer^.ud_Data * 8; // Used-Flag, Modulkennung(SDIAS)
            else
              ud_Address += p_SDOResponseBuffer^.ud_Data * 4; // Used-Flag
            end_if;

          end_if;

//*****************************************************************************
//**   SAFE BOOL INTERFACE OUTPUT VARIABLES                                  **
//*****************************************************************************

          // safe bool interface output vars
          //send request and receive data
          sd_retval := SDOReadCfgRequ ( p_SDORequestBuffer  := p_SDORequestBuffer
                                      , p_SDOResponseBuffer := p_SDOResponseBuffer
                                      , ud_Address          := ud_Address
                                      , us_Length           := 4
                                      );

          //no response
          if ( sd_retval <> 0 ) then
            LogError("@0223 (SafetyBaseFSoE::ReadSDOConfig) Config Read Error: Reading number of safe BOOL interface output variables failed.");
            return;
          end_if;

          // skip safe BOOL interface output variables
          ud_Address += 4;

          // count the interface output variables
          BoolOuts := p_SDOResponseBuffer^.ud_Data;

          if b_IsFSoE then
            ud_TmpCnt := p_SDOResponseBuffer^.ud_Data;

            if ud_TmpCnt then
              for i := 1 to ud_TmpCnt do
                //send request and receive data
                sd_retval := SDOReadCfgRequ ( p_SDORequestBuffer  := p_SDORequestBuffer
                                            , p_SDOResponseBuffer := p_SDOResponseBuffer
                                            , ud_Address          := ud_Address
                                            , us_Length           := 4
                                            );

                //no response
                if ( sd_retval <> 0 ) then
                  LogError("@027A (SafetyBaseFSoE::ReadSDOConfig) Config Read Error: Reading number of FSoE connections for BOOL interface outputs failed.");
                  return;
                end_if;

                // skip number of entries and the entries
                ud_Address += 4 + 4 * p_SDOResponseBuffer^.ud_Data;
              end_for;
            end_if;
          end_if;

//*****************************************************************************
//**   SAFE DINT INTERFACE OUTPUT VARIABLES                                  **
//*****************************************************************************

          // safe dint interface output vars
          //send request and receive data
          sd_retval := SDOReadCfgRequ ( p_SDORequestBuffer  := p_SDORequestBuffer
                                      , p_SDOResponseBuffer := p_SDOResponseBuffer
                                      , ud_Address          := ud_Address
                                      , us_Length           := 4
                                      );

          //no response
          if ( sd_retval <> 0 ) then
            LogError("@0224 (SafetyBaseFSoE::ReadSDOConfig) Config Read Error: Reading number of safe DINT interface output variables failed.");
            return;
          end_if;

          // skip number of safe dint interface output vars
          ud_Address += 4;

          // count the interface output variables
          DintOuts := p_SDOResponseBuffer^.ud_Data;

          if b_IsFSoE then
            ud_TmpCnt := p_SDOResponseBuffer^.ud_Data;

            if ud_TmpCnt then
              for i := 1 to ud_TmpCnt do
                //send request and receive data
                sd_retval := SDOReadCfgRequ ( p_SDORequestBuffer  := p_SDORequestBuffer
                                            , p_SDOResponseBuffer := p_SDOResponseBuffer
                                            , ud_Address          := ud_Address
                                            , us_Length           := 4
                                            );

                //no response
                if ( sd_retval <> 0 ) then
                  LogError("@027B (SafetyBaseFSoE::ReadSDOConfig) Config Read Error: Reading number of FSoE connections for DINT interface outputs failed.");
                  return;
                end_if;

                // skip number of entries and the entries
                ud_Address += 4 + 4 * p_SDOResponseBuffer^.ud_Data;
              end_for;
            end_if;
          end_if;

//*****************************************************************************
//**   FSBs = Functional Safety Blocks                                       **
//*****************************************************************************

          ud_skipLength := 0;

          // skip FSBs! structure: CRC, Length.... until the length is 0
          repeat

            // skip CRC and length of FSB
            ud_Address += 4 + ud_skipLength;

            //send request and receive data
            sd_retval := SDOReadCfgRequ ( p_SDORequestBuffer  := p_SDORequestBuffer
                                        , p_SDOResponseBuffer := p_SDOResponseBuffer
                                        , ud_Address          := ud_Address
                                        , us_Length           := 4
                                        );

            //no response
            if ( sd_retval <> 0 ) then
              LogError("@0225 (SafetyBaseFSoE::ReadSDOConfig) Config Read Error: Reading length of FSB failed.");
              return;
            end_if;

            ud_skipLength := p_SDOResponseBuffer^.ud_Data;

          until ud_skipLength = 0 end_repeat;

          // skip length of block with 0 length
          ud_Address += 4;

          if b_CfgTypeV3 then

//*****************************************************************************
//**   DYNAMIC PARAMETERS (e.g. for SSI Module)                              **
//*****************************************************************************

// Version of Parameters is saved in hd_DynParaVersion
// if it's 16#0001, then we read out the number of parameters which will follow

// structure:
// number of parameters
// for every parameter: place, id, length (including the 4 byte for the length itself), data

            //send request and receive data
            sd_retval := SDOReadCfgRequ ( p_SDORequestBuffer  := p_SDORequestBuffer
                                        , p_SDOResponseBuffer := p_SDOResponseBuffer
                                        , ud_Address          := ud_Address
                                        , us_Length           := 4
                                        );

            //no response
            if ( sd_retval <> 0 ) then
              LogError("@0226 (SafetyBaseFSoE::ReadSDOConfig) Config Read Error: Reading number of dynamic parameters failed.");
              return;
            end_if;

            ud_TmpCnt := p_SDOResponseBuffer^.ud_Data;

            // skip number of parameters
            ud_Address += 4;

            if ud_TmpCnt then
              for i := 1 to ud_TmpCnt do
                //send request and receive data
                sd_retval := SDOReadCfgRequ ( p_SDORequestBuffer  := p_SDORequestBuffer
                                            , p_SDOResponseBuffer := p_SDOResponseBuffer
                                            , ud_Address          := ud_Address
                                            , us_Length           := sizeof(t_DynamicParameterHeader)
                                            );

                //no response
                if ( sd_retval <> 0 ) then
                  LogError("@0227 (SafetyBaseFSoE::ReadSDOConfig) Config Read Error: Reading header of dynamic parameter failed.");
                  return;
                end_if;

                DynamicParameterHeader := p_SDOResponseBuffer^.ud_Data$t_DynamicParameterHeader;

                AddressServiceDataSize := 0;

                // skip size of header
                ud_Address += sizeof(t_DynamicParameterHeader);

                // data for pdo length info:
                // this data is also mirrored to SBF_SDO_ADDRESS_SPECIAL_INFO

//                  Marked with Place = 1000
//
//                  (4 Byte Length)
//                   4 Byte Version (starting at 0)
//                   1 Byte Length Rd PDO
//                   1 Byte Length Rd PDO IF
//                   1 Byte Length Wr PDO
//                   1 Byte Number of write PDOs (without additional it would be 1), msb = fast unsafe active

                if (DynamicParameterHeader.Place = SBF_CONFIG_PDO_INFO_PLACE) & (DynamicParameterHeader.Length >= (sizeof(UDINT) + sizeof(t_PDOSizeInfo))) then
                  //send request and receive data
                  sd_retval := SDOReadCfgRequ ( p_SDORequestBuffer  := p_SDORequestBuffer
                                              , p_SDOResponseBuffer := p_SDOResponseBuffer
                                              , ud_Address          := ud_Address
                                              , us_Length           := sizeof(t_PDOSizeInfo)
                                              );

                  //no response
                  if ( sd_retval <> 0 ) then
                    LogError("@0228 (SafetyBaseFSoE::ReadSDOConfig) Config Read Error: Reading dynamic parameter for pdo size failed.");
                    return;
                  end_if;

                  ud_Address += sizeof(t_PDOSizeInfo);

                  AddressServiceDataSize := (ud_ListLength_Address + ud_ListLength) - ud_Address;

                  PdoSizeInfo := p_SDOResponseBuffer^.ud_Data$t_PDOSizeInfo;

                  //check version
                  if PdoSizeInfo.Version = 1 then
                    // if any sizes increased or we would need more DOs
                    if (PdoSizeInfo.PDORdLen > MyPDOReadSize)     |
                       (PdoSizeInfo.PDOWrLen > MyPDOWriteSize)    |
                       ((PdoSizeInfo.FastUnsafeAvailable <> 0) > ActivateFastUnsafeIOs) then

                      // error => can't go on like this
                      LogError("@0202 (SafetyBaseFSoE::ReadSDOConfig) Number or size of module accesses increased with new safety project!");
                      LogError("@0203 (SafetyBaseFSoE::ReadSDOConfig) => Can't continue, because the new data is not covered by the actual accesses! Restart Application!");

                      b_NeedApplicationRestart := TRUE;
                    end_if;
                  else
                    // new interpretercode version
                    PdoSizeInfoV2 := p_SDOResponseBuffer^.ud_Data$t_PDOSizeInfoV2;

                    if  (PdoSizeInfoV2.PDORdLen > MyPDOReadSize)                       |
                        (PdoSizeInfoV2.PDOWrLen > MyPDOWriteSize)                      |
                        (PdoSizeInfoV2.uiNumberFastUnsafeRdVar > uiNumberFastUnsafeRd) |
                        (PdoSizeInfoV2.uiNumberFastUnsafeWrVar > uiNumberFastUnsafeWr) then

                      // error => can't go on like this
                      LogError("@0202 (SafetyBaseFSoE::ReadSDOConfig) Number or size of module accesses increased with new safety project!");
                      LogError("@0203 (SafetyBaseFSoE::ReadSDOConfig) => Can't continue, because the new data is not covered by the actual accesses! Restart Application!");

                      b_NeedApplicationRestart := TRUE;
                    end_if;
                  end_if;

                  exit;
                end_if;

                // skip the parameter data (length of the length is also included)
                ud_Address += DynamicParameterHeader.Length - 4;
              end_for;

              if AddressServiceDataSize then
(*

  Data structure of address service data

  4 Byte Anzahl der MultiChannel
    Pro MultiChannel:
    4 Byte Anzahl der Verwendungen des Multichannel
    4 Byte Index des Gesamtergebnisses
    1 Byte Art der Verknüpfung (0 = UND)
    1 Byte Defaultbelegung des Werts
    2 Byte Reserved (für 4 Byte Alignment)
      Pro Verwendung (siehe erster Eintrag in den MultiChannelDaten):
      4 Byte FSoE Daten
  4 Byte Kommunikations-ID (Default 0)
  4 Byte Anzahl der Adressbereiche
    Pro Adressbereich:
    4 Byte Startadresse
    4 Byte Länge Adressbereich
  4 Byte Anzahl der Connection-ID-Bereiche
    Pro Bereich:
    4 Byte Startadresse
    4 Byte Länge Bereich

*)
                // get the number of multichannels
                sd_retval := SDOReadCfgRequ ( p_SDORequestBuffer  := p_SDORequestBuffer
                                            , p_SDOResponseBuffer := p_SDOResponseBuffer
                                            , ud_Address          := ud_Address
                                            , us_Length           := 4
                                            );

                //no response
                if ( sd_retval <> 0 ) then
                  LogError("@027C (SafetyBaseFSoE::ReadSDOConfig) Config Read Error: Reading address service data failed.");
                  return;
                end_if;

                ud_TmpCnt := p_SDOResponseBuffer^.ud_Data;

                // skip number of multichannels
                ud_Address += 4;

                if ud_TmpCnt then
                  for i := 1 to ud_TmpCnt do
                    // get the number of usages
                    sd_retval := SDOReadCfgRequ ( p_SDORequestBuffer  := p_SDORequestBuffer
                                                , p_SDOResponseBuffer := p_SDOResponseBuffer
                                                , ud_Address          := ud_Address
                                                , us_Length           := 4
                                                );

                    //no response
                    if ( sd_retval <> 0 ) then
                      LogError("@027C (SafetyBaseFSoE::ReadSDOConfig) Config Read Error: Reading address service data failed.");
                      return;
                    end_if;

                    // skip the rest of this multichannel
                    ud_Address += 12 + (p_SDOResponseBuffer^.ud_Data * 4);
                  end_for;
                end_if;

                // skip the communication ID
                ud_Address += 4;

                // read the number of address areas
                sd_retval := SDOReadCfgRequ ( p_SDORequestBuffer  := p_SDORequestBuffer
                                            , p_SDOResponseBuffer := p_SDOResponseBuffer
                                            , ud_Address          := ud_Address
                                            , us_Length           := 4
                                            );

                //no response
                if ( sd_retval <> 0 ) then
                  LogError("@027C (SafetyBaseFSoE::ReadSDOConfig) Config Read Error: Reading address service data failed.");
                  return;
                end_if;

                // if there are any => the module got an address service
                if p_SDOResponseBuffer^.ud_Data then
                  TempModuleConfig.Info.IsAddressService := TRUE;
                end_if;
              end_if;
            end_if;
          end_if;

          // if there are interface variables
          if BoolOuts | DintOuts then
            // calculate the length of the interface frame
            TempPdoConfig.PdoLen := CalcPDOLength(BoolOuts, DintOuts);

            TempPdoConfig.Info := 0;
            TempPdoConfig.Info.IsInterfacePDO := TRUE;
            TempPdoConfig.Info.IsOptional := (ud_ActBlockType = SBF_BLKTYPE_CFG_MODULE_OPTIONAL);

            // if it's a broadcast => mark it
            if (TempPath[0]$UINT = 2) & (TempPath[0]$HDINT = SBF_INTERFACE_FRAME_BROADCAST) then
              TempPdoConfig.Info.IFBroadCast := TRUE;
            end_if;

            // this is the source of the interface frame
            TempPdoConfig.SourcePathLen := pListHeader^.p_us_Path^$UINT + 2;
            TempPdoConfig.pSourcePath   := pListHeader^.p_us_Path;

            // and the destination
            TempPdoConfig.DestPathLen   := TempPath[0]$UINT + 2;
            TempPdoConfig.pDestPath     := #TempPath[0];

            // add the interface PDO to the list
//            AddPdoToCfg(TempPdoConfig);

            TempModuleConfig.Info.IsInterfaceSource := TRUE;
            TempModuleConfig.Info.IsInterfaceDest   := FALSE;
            TempModuleConfig.InterfaceCRC := TempPdoConfig.InterfaceCRC;
          else
            TempModuleConfig.Info.IsInterfaceSource := FALSE;
            TempModuleConfig.Info.IsInterfaceDest   := FALSE;
            TempModuleConfig.InterfaceCRC := 0;
          end_if;
        else
          TempModuleConfig.Info.IsInterfaceSource := FALSE;
          TempModuleConfig.Info.IsInterfaceDest   := FALSE;
          TempModuleConfig.InterfaceCRC := 0;
        end_if;

        // if it's our own path, remember the safety number
        if (PathOfThisCPU[0]$UINT = (pListHeader^.p_us_Path$^UINT)^) & (ToStdLib.MemCmp(#PathOfThisCPU[0], pListHeader^.p_us_Path, PathOfThisCPU[0]$UINT + 2) = 0) then
          TempModuleConfig.SafetyNbr := SafetyNumber;
          //safe config of scp modul (own path)
          SafeActModuleConfig(TempModuleConfig);
        else
          TempModuleConfig.SafetyNbr := 0;
        end_if;

        // only when there is a manager
        if pSafetyManagerThis then
          AddModuleToCfg(TempModuleConfig);
        end_if;

//**********************************************************************************************************************************************************
      SBF_BLKTYPE_OLD_MODE_FLAG: // flag fore FW to use old config-mode
        // we need the old TimeSync config-type
        NewConfigType := ConfigState_Old;

//**********************************************************************************************************************************************************
      SBF_BLKTYPE_CFG_XML: // configuration for uploading the project to the safetydesigner (network placement information, names of bits,...)
        // no useful information here for us

//**********************************************************************************************************************************************************
    else
      // skip it = do nothing
//      TRACE("Found unhandled Blocktype in configuration.");
//**********************************************************************************************************************************************************
    end_case;

    ud_ListBaseAddress := ud_ListLength_Address + ud_ListLength;
  end_while;

  if ( ( sd_retval = 0 ) & ( SafetyState = _ModFromCfgNotFound ) ) then
    sd_retval := -1;
  end_if;

END_FUNCTION

FUNCTION VIRTUAL SafetyBaseFSoE::SDOReadCfgRequ
  VAR_INPUT
    p_SDORequestBuffer 	: ^SafetyBaseFSoE::SDORequReadConfig;
    p_SDOResponseBuffer 	: ^SafetyBaseFSoE::SDORespReadConfig;
    ud_Address 	: UDINT;
    us_Length 	: USINT;
    b_UseCache 	: BOOL;(* := TRUE *)
  END_VAR
  VAR_OUTPUT
    sd_retval 	: DINT;
  END_VAR

  // check if we have the data in the cache
  if b_UseCache & IsInCache(ud_Address, us_Length) then
    // use it from the cache

    // the address may be used from outside this function
    p_SDORequestBuffer^.ud_Address := ud_Address;

    _memcpy(ptr1:=#p_SDOResponseBuffer^.ud_Data, ptr2:=#Cache[0] + (ud_Address - CachedAddr), cntr:=us_Length);

    // everything is fine
    sd_retval := 0;
  else

    //sequence number
    p_SDORequestBuffer^.StdHeader.SeqNr := us_CntSequNr;

    //increase counter for sequence number
    if us_CntSequNr < 16#7F then
      us_CntSequNr += 1;
    else
      us_CntSequNr := 0;
    end_if;

    //address
    p_SDORequestBuffer^.ud_Address := ud_Address;

    if b_UseCache then
      // get max size
      p_SDORequestBuffer^.us_Length := SBF_SDO_MAX_LENGTH - (sizeof(SDORespReadConfig) - sizeof(SDORespReadConfig.ud_Data));
    else
      //length of expected data
      p_SDORequestBuffer^.us_Length := us_Length;
    end_if;

    //calculate CRC (starting with length of data until the end of command)
    p_SDORequestBuffer^.StdHeader.CRC := 0;

    //send request
    sd_retval := SAFETY_iSendRequest( uiMaster    := 0
                                    , pucNode     := p_ObjectPath
                                    , uiInLength  := sizeof(SDORequReadConfig)
                                    , pucInput    := p_SDORequestBuffer$^USINT
                                    , uiOutLength := sizeof(SDORespReadConfig) - sizeof(SDORespReadConfig.ud_Data) + p_SDORequestBuffer^.us_Length
                                    , pucOutput   := p_SDOResponseBuffer$^USINT
                                    );

    //no response
    if ( sd_retval <> 0 ) then
      LogError("@0229 (SafetyBaseFSoE::SDOReadCfgRequ) SAFETY_iSendRequest failed.");

      // we remember to retry in a few seconds
      b_ReadConfigFailed := TRUE;
      return;
    end_if;

    //check sequence number to exclude a possible wrong response
    if ( p_SDORequestBuffer^.StdHeader.SeqNr <> p_SDOResponseBuffer^.StdHeader.SeqNr ) then
      // we remember to retry in a few seconds
      b_ReadConfigFailed := TRUE;
      //log not routable SDOs
      LogValue("@022A (SafetyBaseFSoE::SDOReadCfgRequ) Invalid Sequence number in SDO Standard Response. Got 0x{0} instead of expected 0x{1}", to_udint(p_SDOResponseBuffer^.StdHeader.SeqNr), to_udint(p_SDORequestBuffer^.StdHeader.SeqNr));
      return;
    end_if;

    //check returncode of SDO
    if ( p_SDOResponseBuffer^.us_Returncode <> SBF_SDO_RETCODE_OK ) then
      //log not routable SDOs
      LogValue("@022B (SafetyBaseFSoE::SDOReadCfgRequ) Safety module 0x{0}: Retcode of SDO Standard Response was invalid. Retcode: 0x{1}", SafetyNumber$UDINT, to_udint(p_SDOResponseBuffer^.us_Returncode));

  //    // when reading fails because safety designer is writing at the same moment
  //    if p_SDOResponseBuffer^.us_Returncode = SDO_MICROCTRL_DIFFER then
        // we remember to retry in a few seconds
        b_ReadConfigFailed := TRUE;
  //    end_if;

      return;
    end_if;

    //check length of read data
    if ( p_SDOResponseBuffer^.us_Length = 0 ) then
      LogError("@022C (SafetyBaseFSoE::SDOReadCfgRequ) Response length is 0.");
      sd_retval := -104;
      return;
    elsif b_UseCache then
      // everything is fine => add the new data to the cache
      AddToCache(p_SDORequestBuffer, p_SDOResponseBuffer);
    end_if;
  end_if;

END_FUNCTION

FUNCTION VIRTUAL SafetyBaseFSoE::GetRoutingData
  VAR_OUTPUT
    sd_retval 	: DINT;
  END_VAR
  VAR
    SDORequestBuffer        : SDORequReadConfig;
    SDOResponseBuffer       : ARRAY [0..SBF_SDO_MAX_LENGTH-1] OF USINT;
    p_SDORequestBuffer 	    : ^SDORequReadConfig;
    p_SDOResponseBuffer 	  : ^SDORespReadConfig;
    Module                  : PathInfoType;
    ListHeader              : PathInfoType;
    NotAvailableStr         : ARRAY [0..99] OF CHAR;
    ModulePath              : ARRAY [0..127] OF USINT;
    ModulePathComp          : ARRAY [0..127] OF USINT;
    ListPath                : ARRAY [0..127] OF USINT;
    ListPathComp            : ARRAY [0..127] OF USINT;
    Time1, Time2            : UDINT;
  END_VAR

  // get module specific configuration information
  GetConfiguration();

  InitPathInfo(#Module);
  InitPathInfo(#ListHeader);

  //SDO request for this command has 5 bytes additional to the header
  p_SDORequestBuffer := #SDORequestBuffer;

  //SDO response for this command can have maximum additional data
  p_SDOResponseBuffer := (#SDOResponseBuffer)$^SDORespReadConfig;

  //path of input-safety-module
  Module.p_us_Path$^void := #ModulePath;

  //compressed path of input-safety-module
  Module.p_us_PathComp$^void := #ModulePathComp;

  //path in list header
  ListHeader.p_us_Path$^void := #ListPath;

  //path in list header
  ListHeader.p_us_PathComp$^void := #ListPathComp;

  repeat
    // if not used => continue
    // if valid    => set to not used and continue
    // if wait4rt  => wait in the loop until the state changes to valid
  until (sigclib_atomic_cmpxchgU32(pValue:=#udConfigValid, cmpVal:=SBF_LOCKCFG_VALID, newVal:=SBF_LOCKCFG_NOT_USED) < SBF_LOCKCFG_WAIT4RT) end_repeat;

  b_ReadConfigFailed := FALSE;

  b_NeedApplicationRestart := FALSE;

  // if there is a revision in the configuration this variable changes to TRUE
  b_GotNewRevision := FALSE;

Time1 := OS_READMICROSEC();
  //read config data via SDOs and add safety modules to routing lists
  sd_retval := ReadSDOConfig( p_SDORequestBuffer      := p_SDORequestBuffer
                            , p_SDOResponseBuffer     := p_SDOResponseBuffer
                            , pModule                 := #Module
                            , pListHeader             := #ListHeader
                            );
Time2 := OS_READMICROSEC();
ud_ConfigReadTime := Time2 - Time1;

  // set error to restart application afterwards to have a complete configuration (needed for routing to share the slave configurations with only 1 restart of the application)
  if b_NeedApplicationRestart then
    SetSafetyState(NewState:=_DOsIncreasedRestartApp);
    b_GetNewConfiguration := FALSE; // don't try again (unless the CRC changes again)
    sd_retval := -1;
  end_if;

  // if there is no revision in the configuration => clear it
  if (b_GotNewRevision = FALSE) then

    // free memory, if available
    if pPrjNameStr & pPrjRevStr then
      ToStdLib.Free(pPrjNameStr);
    end_if;

    // use local memory to show "not available"
    _strcpy(dest:=#NotAvailableStr[0], src:="<not available>");
    PrjNameMemLen := _strlen(src:=#NotAvailableStr[0]);
    PrjNameStrLen := PrjRevStrLen := PrjNameMemLen - 1;
    pPrjNameStr := pPrjRevStr := #NotAvailableStr[0];

    // write the strings to the string objects
    ShowProjectRevision();

    // there is no memory, so reset the pointer and length informations
    pPrjNameStr := NIL;
    pPrjRevStr := NIL;

    PrjNameMemLen := 0;
    PrjNameStrLen := 0;
    PrjRevStrLen := 0;
  end_if;

  // if reading failed, because designer is writing at the same time => we try again in a few seconds
  if b_ReadConfigFailed then

    // next time we check for the configured state of the cpu
    b_CheckConfigured := TRUE;
    b_GetNewConfiguration := FALSE; // don't try again while the config is invalid

    // check again in background
    SetSafetyState(NewState:=_ReinitConfig);

    // and wait at least 3 secs
    ud_LastCheckConfig := ops.tAbsolute;

  // error in configuration -> no work
  elsif ( sd_retval <> 0 ) & (SafetyState <> _ReinitConfig) then
    if SafetyState = _WaitForSynchronicity then
      SetSafetyState(NewState:=_UnknownCfgError);
    end_if;

    LogError("@022D (SafetyBaseFSoE::GetRoutingData) Reading Safety Configuration failed!");
  else
    // read config succeeded, check update cycle of unsafe variables
    CheckUnsafeUpdateCycle();

    // check for interface frame destination modules and mark them
    GetDestinationCRCs();

    // if there is a safety manager create a configuration message and send it to the safety manager
    if pSafetyManagerThis then
      CreateAndSendCfg();
    end_if;

    // last thing to do is to start realtime and cyclic work (they do nothing in _ReinitConfig state)
    if ud_UnsafeVarsNotFound then
      SetSafetyState(NewState:=_UnsafeVarNotFound);
      ud_UnsafeVarsNotFound := 0;
    else
      if us_SetBusReadyState = SetBusReadyFinished then
        // we're already synchron from a former configuration phase
        SetSafetyState(NewState:=_SafetyClassOK);
      else
        SetSafetyState(NewState:=_WaitForSynchronicity);
      end_if;
    end_if;

    // set config valid
    sigclib_atomic_swpU32(pValue:=#udConfigValid, swpVal:=SBF_LOCKCFG_VALID);
  end_if;

  // free temporary configuration lists if there were any
  FreeCfgLists();

END_FUNCTION

FUNCTION VIRTUAL SafetyBaseFSoE::ReadModulePath
  VAR_INPUT
    p_SDORequestBuffer 	: ^SafetyBaseFSoE::SDORequReadConfig;
    p_SDOResponseBuffer 	: ^SafetyBaseFSoE::SDORespReadConfig;
    p_ud_Address 	: ^UDINT;
    pModule 	: ^SafetyBaseFSoE::PathInfoType;
    p_ud_ModulePathLen_Max 	: ^UDINT;
    p_ud_ModulePathCompLen_Max 	: ^UDINT;
    us_SDOMaxDataSize 	: USINT;
  END_VAR
  VAR_OUTPUT
    sd_retval 	: DINT;
  END_VAR
  VAR
    ud_ModulePathLen_Act    : UDINT;
    p_ud_ModulePath_Act     : ^UDINT;
  END_VAR

  //read length of module path

  //send request and receive data
  sd_retval := SDOReadCfgRequ ( p_SDORequestBuffer  := p_SDORequestBuffer
                              , p_SDOResponseBuffer := p_SDOResponseBuffer
                              , ud_Address          := p_ud_Address^
                              , us_Length           := 4
                              );

  //no response
  if ( sd_retval <> 0 ) then
    LogError("@022E (SafetyBaseFSoE::ReadModulePath) Failed to read length of module path.");
    return;
  end_if;

  //length of module path
  ud_ModulePathLen_Act := p_SDOResponseBuffer^.ud_Data;

  //length is zero, check compressed path
  if ( ud_ModulePathLen_Act > 0 ) then

    // if it's too small => error
    if ( ud_ModulePathLen_Act > p_ud_ModulePathLen_Max^ ) then
      sd_retval                         := -100;
      SetSafetyState(NewState:=_MemAllocFailed);
      return;
    end_if;

    //read path

    //address of first byte of path
    p_ud_Address^ += 4;

    //set pointer to first byte of target buffer
    p_ud_ModulePath_Act := ( pModule^.p_us_Path )$^UDINT;

    //read path block by block, if path is longer than max. length
    while ( ud_ModulePathLen_Act > us_SDOMaxDataSize ) do

      //send request and receive data
      sd_retval := SDOReadCfgRequ ( p_SDORequestBuffer  := p_SDORequestBuffer
                                  , p_SDOResponseBuffer := p_SDOResponseBuffer
                                  , ud_Address          := p_ud_Address^
                                  , us_Length           := us_SDOMaxDataSize
                                  , b_UseCache          := FALSE
                                  );

      //no response
      if ( sd_retval <> 0 ) then
        LogError("@022F (SafetyBaseFSoE::ReadModulePath) Failed to read block of module path.");
        return;
      end_if;

      //copy part of path
      ToStdLib.MemCpy(dest := p_ud_ModulePath_Act , source := #p_SDOResponseBuffer^.ud_Data, size := us_SDOMaxDataSize);

      //rest of path to be read
      ud_ModulePathLen_Act -= us_SDOMaxDataSize;

      //address of next block
      p_ud_Address^ += us_SDOMaxDataSize;

      //set pointer to next free byte of target buffer
      p_ud_ModulePath_Act += us_SDOMaxDataSize;

    end_while;

    // if there is something left
    if ud_ModulePathLen_Act then
      //read last bytes of path

      //send request and receive data
      sd_retval := SDOReadCfgRequ ( p_SDORequestBuffer  := p_SDORequestBuffer
                                  , p_SDOResponseBuffer := p_SDOResponseBuffer
                                  , ud_Address          := p_ud_Address^
                                  , us_Length           := ud_ModulePathLen_Act$USINT
                                  , b_UseCache          := ud_ModulePathLen_Act$USINT < us_SDOMaxDataSize
                                  );

      //no response
      if ( sd_retval <> 0 ) then
        LogError("@0230 (SafetyBaseFSoE::ReadModulePath) Failed to read last bytes of module path.");
        return;
      end_if;

      ToStdLib.MemCpy(dest := p_ud_ModulePath_Act, source := #p_SDOResponseBuffer^.ud_Data, size := ud_ModulePathLen_Act);
    end_if;
